Fanuc KAREL source: KT00671.KL

PROGRAM KT00671
%NOLOCKGROUP
VAR
  P1: XYZWPREXT
  P2: XYZWPREXT
  OUT: REAL
BEGIN
  P1.X = 1.0
  P2.Y = 2.0
  P1.X = 1.0
  P2.Y = 2.0
  OUT = NOT P1
END KT00671
